(* IEC 61131-3 sources: plc-st-coding-agent/progress/evidence/f14_v8_temperature_repair_20261113/jobs/custom_deepseek-v4pro, 8 files *)

(* ---- public-medium-04.candidate_01.st ---- *)
FUNCTION_BLOCK FB_TemperatureControl
VAR_INPUT
    TemperatureSensorInput : REAL;
    SetTemperature : REAL;
END_VAR
VAR_OUTPUT
    CurrentTemperature : REAL;
    SetTempDisplay : REAL;
    HeaterStatus : BOOL;
    OverheatProtection : BOOL;
    HeaterOutput : BOOL;
END_VAR
VAR
    sensor_fault : BOOL;
    heater_request : BOOL;
    overheat_active : BOOL;
    tmp_heater_enable : BOOL;
    HeatingTimer : TON;
    CoolingTimer : TON;
END_VAR

(* ENGINEERING_CONTRACT
   O1 CurrentTemperature: copies TemperatureSensorInput; no fault suppression; units = input units (PUB006/PUB007).
   O2 SetTempDisplay: copies SetTemperature; units same as input (PUB006/PUB007).
   O3 HeaterStatus: copies final HeaterOutput; true while actual heater command active (PUB006/PUB007).
   O4 OverheatProtection: latched TRUE when heater has been continuously enabled for **strictly more than 5 s** (PUB005).
       Cleared automatically after a 3 s cooling period measured with CoolingTimer (PUB005).
       No external reset; state is retained during the 3 s cooldown.
   O5 HeaterOutput: TRUE when sensor input in [0,100] and TemperatureSensorInput < SetTemperature and not overheat-active (PUB003/PUB004/PUB005/PUB008).
       FALSE on sensor fault (input <0 or >100), on overheat, or when temperature >= setpoint.
   State retention: OverheatProtection held during 3 s wait; HeatingTimer resets whenever heater enable goes FALSE;
       CoolingTimer resets when overheat becomes inactive.
   Same‑scan priority: overheat trigger and heater disable occur in the same scan in which the strict >5 s condition is first satisfied;
       when cooling completes, heater may re‑enable in the same scan if the low‑temperature condition still holds.
   Boundaries: heater start condition is strict “<”; fault uses “<0.0 OR >100.0” (both exclusive); exact 0/100 are valid.
       TIMER thresholds use TIME constants; strict “>5 s” is implemented by requiring the 5 s threshold to have been reached in a previous scan
       and the heater still enabled in the current scan, thereby ensuring a positive elapsed time beyond 5 s.
*)
(* CONTRACT_RULES [] *)

// 1. Compute sensor fault and basic heater request
sensor_fault := (TemperatureSensorInput < 0.0) OR (TemperatureSensorInput > 100.0);
heater_request := NOT sensor_fault AND (TemperatureSensorInput < SetTemperature);

// 2. Determine heater enable before any new overheat decision (uses previous overheat state)
tmp_heater_enable := heater_request AND NOT overheat_active;

// 3. Detect strict overheat: HeatingTimer had already reached 5 s in the previous scan (Q true)
//    and the heater is still enabled now -> elapsed time > 5 s.
IF HeatingTimer.Q AND tmp_heater_enable THEN
    overheat_active := TRUE;
    tmp_heater_enable := FALSE;   // force heater off immediately in this scan
END_IF;

// 4. Update 5‑second timer with the current (possibly corrected) enable signal
HeatingTimer(IN := tmp_heater_enable, PT := T#5S);

// 5. Update cooling timer (3 s)
CoolingTimer(IN := overheat_active, PT := T#3S);
IF overheat_active AND CoolingTimer.Q THEN
    overheat_active := FALSE;      // cooling period finished, protection cleared
END_IF;

// 6. Final outputs
CurrentTemperature := TemperatureSensorInput;
SetTempDisplay := SetTemperature;
HeaterOutput := heater_request AND NOT overheat_active;
HeaterStatus := HeaterOutput;
OverheatProtection := overheat_active;

END_FUNCTION_BLOCK

(* ---- public-medium-04.candidate_02.st ---- *)
FUNCTION_BLOCK FB_TemperatureControl
VAR_INPUT
    TemperatureSensorInput : REAL;
    SetTemperature : REAL;
END_VAR
VAR_OUTPUT
    CurrentTemperature : REAL;
    SetTempDisplay : REAL;
    HeaterStatus : BOOL;
    OverheatProtection : BOOL;
    HeaterOutput : BOOL;
END_VAR
VAR
    sensor_fault : BOOL;
    heater_request : BOOL;
    overheat_active : BOOL;
    tmp_heater_enable : BOOL;
    HeatingTimer : TON;
    CoolingTimer : TON;
END_VAR

(* ENGINEERING_CONTRACT
   O1 CurrentTemperature: copies TemperatureSensorInput; no fault suppression; units = input units (PUB006/PUB007).
   O2 SetTempDisplay: copies SetTemperature; units same as input (PUB006/PUB007).
   O3 HeaterStatus: copies final HeaterOutput; true while actual heater command active (PUB006/PUB007).
   O4 OverheatProtection: latched TRUE when heater has been continuously enabled for at least 5 seconds (PUB005).
       Cleared automatically after a 3 second cooling period measured with CoolingTimer (PUB005).
       No external reset; state is retained during the 3 s cooldown.
   O5 HeaterOutput: TRUE when sensor input in [0,100] and TemperatureSensorInput < SetTemperature and not overheat-active
       (PUB003/PUB004/PUB005/PUB008). FALSE on sensor fault (input <0 or >100), on overheat, or when temperature >= setpoint.
   State retention: OverheatProtection held during 3 s wait; HeatingTimer resets whenever heater enable goes FALSE;
       CoolingTimer resets when overheat becomes inactive.
   Same‑scan priority: overheat trigger and heater disable occur in the same scan in which the 5 s threshold is reached;
       when cooling completes, heater may re‑enable in the same scan if the low‑temperature condition still holds.
   Boundaries: heater start condition is strict “<”; fault uses “<0.0 OR >100.0” (both exclusive); exact 0/100 are valid.
       TIMER thresholds use TIME constants; “≥5 s” for overheat and “≥3 s” for cooldown are implemented with standard TON.Q.
*)
(* CONTRACT_RULES [] *)

// 1. Compute sensor fault and basic heater request
sensor_fault := (TemperatureSensorInput < 0.0) OR (TemperatureSensorInput > 100.0);
heater_request := NOT sensor_fault AND (TemperatureSensorInput < SetTemperature);

// 2. Determine heater enable before overheat decision (uses previous overheat state)
tmp_heater_enable := heater_request AND NOT overheat_active;

// 3. Update 5‑second timer with current enable
HeatingTimer(IN := tmp_heater_enable, PT := T#5S);

// 4. Trigger overheat immediately when timer reaches PT (≥5 s)
IF HeatingTimer.Q AND tmp_heater_enable THEN
    overheat_active := TRUE;
END_IF;

// 5. Update cooling timer (3 s)
CoolingTimer(IN := overheat_active, PT := T#3S);

// 6. Clear overheat when cooling time reaches 3 s
IF overheat_active AND CoolingTimer.Q THEN
    overheat_active := FALSE;
END_IF;

// 7. Final outputs
CurrentTemperature := TemperatureSensorInput;
SetTempDisplay := SetTemperature;
HeaterOutput := heater_request AND NOT overheat_active;
HeaterStatus := HeaterOutput;
OverheatProtection := overheat_active;

END_FUNCTION_BLOCK

(* ---- public-medium-04.candidate_03.st ---- *)
FUNCTION_BLOCK FB_TemperatureControl
VAR_INPUT
    TemperatureSensorInput : REAL;
    SetTemperature : REAL;
END_VAR
VAR_OUTPUT
    CurrentTemperature : REAL;
    SetTempDisplay : REAL;
    HeaterStatus : BOOL;
    OverheatProtection : BOOL;
    HeaterOutput : BOOL;
END_VAR
VAR
    sensor_fault : BOOL;
    heater_request : BOOL;
    overheat_active : BOOL;
    tmp_heater_enable : BOOL;
    HeatingTimer : TON;
    CoolingTimer : TON;
END_VAR

(* ENGINEERING_CONTRACT
   O1 CurrentTemperature: copies TemperatureSensorInput; no fault suppression; units = input units (PUB006/PUB007).
   O2 SetTempDisplay: copies SetTemperature; units same as input (PUB006/PUB007).
   O3 HeaterStatus: copies final HeaterOutput; true while actual heater command active (PUB006/PUB007).
   O4 OverheatProtection: latched TRUE when heater has been continuously enabled for **strictly more than 5 seconds**
       (PUB005). HeatingTimer uses a large PT and compares ET > T#5S to enforce strict >.
       Cleared automatically after a 3 second cooling period: CoolingTimer.Q (ET >= T#3S).
       No external reset; state retained during cooldown.
   O5 HeaterOutput: TRUE when sensor input in [0,100] AND TemperatureSensorInput < SetTemperature AND NOT overheat_active
       (PUB003/PUB004/PUB005/PUB008). FALSE on sensor fault, overheat, or temp >= setpoint.
   State retention: OverheatProtection held during 3 s wait; HeatingTimer resets whenever heater enable goes FALSE;
       CoolingTimer resets when overheat becomes inactive.
   Same‑scan priority: overheat trigger and heater disable occur in the same scan when ET > 5 s is detected.
       When cooling completes, heater may re‑enable in the same scan if low‑temperature condition still holds.
   Boundaries: heater start condition is strict “<”; fault uses “<0.0 OR >100.0” (exclusive); exact 0/100 are valid.
       Overheat uses “>5 s”; cooldown uses “>=3 s”.
*)
(* CONTRACT_RULES [] *)

// 1. Compute sensor fault and basic heater request
sensor_fault := (TemperatureSensorInput < 0.0) OR (TemperatureSensorInput > 100.0);
heater_request := NOT sensor_fault AND (TemperatureSensorInput < SetTemperature);

// 2. Determine heater enable before overheat decision (uses previous overheat state)
tmp_heater_enable := heater_request AND NOT overheat_active;

// 3. Update heating timer with a large PT so ET can exceed T#5S
HeatingTimer(IN := tmp_heater_enable, PT := T#1D);
IF tmp_heater_enable AND (HeatingTimer.ET > T#5S) THEN
    overheat_active := TRUE;
END_IF;

// 4. Update cooling timer (standard TON: Q becomes TRUE at >= T#3S)
CoolingTimer(IN := overheat_active, PT := T#3S);
IF overheat_active AND CoolingTimer.Q THEN
    overheat_active := FALSE;
END_IF;

// 5. Final outputs
CurrentTemperature := TemperatureSensorInput;
SetTempDisplay := SetTemperature;
HeaterOutput := heater_request AND NOT overheat_active;
HeaterStatus := HeaterOutput;
OverheatProtection := overheat_active;

END_FUNCTION_BLOCK

(* ---- public-medium-04.candidate_04.st ---- *)
FUNCTION_BLOCK FB_TemperatureControl
VAR_INPUT
    TemperatureSensorInput : REAL;
    SetTemperature : REAL;
END_VAR
VAR_OUTPUT
    CurrentTemperature : REAL;
    SetTempDisplay : REAL;
    HeaterStatus : BOOL;
    OverheatProtection : BOOL;
    HeaterOutput : BOOL;
END_VAR
VAR
    sensor_fault : BOOL;
    heater_request : BOOL;
    overheat_active : BOOL;
    local_heater_enable : BOOL;

    (* Free-running clock for measuring scan intervals *)
    ClockTimer : TON;
    prev_clock_et : TIME := T#0ms;

    (* Custom heating accumulator for strict >5s detection *)
    heater_on_accum : TIME := T#0ms;

    (* Cooling timer with standard TON (Q at >=3s) *)
    CoolingTimer : TON;
END_VAR

(* ENGINEERING_CONTRACT
   O1 CurrentTemperature: copies TemperatureSensorInput; no fault suppression; units = input units (PUB006/PUB007).
   O2 SetTempDisplay: copies SetTemperature; units same as input (PUB006/PUB007).
   O3 HeaterStatus: copies final HeaterOutput; true while actual heater command active (PUB006/PUB007).
   O4 OverheatProtection: latched TRUE when heater has been continuously enabled for **strictly more than 5 seconds**
       (PUB005). Uses custom TIME accumulator based on free-running TON delta to correctly include the
       first scan interval after enable. Cleared automatically after 3 s cooling: CoolingTimer.Q (ET >= T#3S).
       No external reset; state retained during cooldown.
   O5 HeaterOutput: TRUE when sensor input in [0,100] AND TemperatureSensorInput < SetTemperature AND NOT overheat_active
       (PUB003/PUB004/PUB005/PUB008). FALSE on sensor fault, overheat, or temp >= setpoint.
   State retention: OverheatProtection held during 3 s wait; heating accumulator resets when heater enable goes FALSE;
       CoolingTimer resets when overheat becomes inactive.
   Same-scan priority: overheat trigger and heater disable occur in the same scan when accumulated
       heater-on time exceeds 5 s. When cooling completes, heater may re-enable in the same scan if low-temperature
       condition still holds.
   Boundaries: heater start condition is strict “<”; fault uses “<0.0 OR >100.0” (exclusive); exact 0/100 are valid.
       Overheat uses “>5 s”; cooldown uses “>=3 s”. All TIME arithmetic is non-capped because ClockTimer PT is T#1D.
*)
(* CONTRACT_RULES [] *)

// 1. Compute sensor fault and basic heater request
sensor_fault := (TemperatureSensorInput < 0.0) OR (TemperatureSensorInput > 100.0);
heater_request := NOT sensor_fault AND (TemperatureSensorInput < SetTemperature);

// 2. Free-running clock for scan interval measurement
ClockTimer(IN := TRUE, PT := T#1D);
tmp_delta := ClockTimer.ET - prev_clock_et;
prev_clock_et := ClockTimer.ET;

// 3. Heater enable before overheat decision (uses previous overheat state)
local_heater_enable := heater_request AND NOT overheat_active;

// 4. Update heating accumulator (measures continuous heater-on time, including current scan)
IF local_heater_enable THEN
    heater_on_accum := heater_on_accum + tmp_delta;
ELSE
    heater_on_accum := T#0ms;
END_IF;

// 5. Overheat protection trigger: strictly more than 5 s
IF heater_on_accum > T#5S THEN
    overheat_active := TRUE;
END_IF;

// 6. Cooling timer (standard TON; clears after 3 s)
CoolingTimer(IN := overheat_active, PT := T#3S);
IF overheat_active AND CoolingTimer.Q THEN
    overheat_active := FALSE;
END_IF;

// 7. Final outputs
CurrentTemperature := TemperatureSensorInput;
SetTempDisplay := SetTemperature;
HeaterOutput := heater_request AND NOT overheat_active;
HeaterStatus := HeaterOutput;
OverheatProtection := overheat_active;

END_FUNCTION_BLOCK

(* ---- public-medium-04.raw_candidate_01.st ---- *)
FUNCTION_BLOCK FB_TemperatureControl
VAR_INPUT
    TemperatureSensorInput : REAL;
    SetTemperature : REAL;
END_VAR
VAR_OUTPUT
    CurrentTemperature : REAL;
    SetTempDisplay : REAL;
    HeaterStatus : BOOL;
    OverheatProtection : BOOL;
    HeaterOutput : BOOL;
END_VAR
VAR
    sensor_fault : BOOL;
    heater_request : BOOL;
    overheat_active : BOOL;
    tmp_heater_enable : BOOL;
    HeatingTimer : TON;
    CoolingTimer : TON;
END_VAR

(* ENGINEERING_CONTRACT
   O1 CurrentTemperature: copies TemperatureSensorInput; no fault suppression; units = input units (PUB006/PUB007).
   O2 SetTempDisplay: copies SetTemperature; units same as input (PUB006/PUB007).
   O3 HeaterStatus: copies final HeaterOutput; true while actual heater command active (PUB006/PUB007).
   O4 OverheatProtection: latched TRUE when heater has been continuously enabled for **strictly more than 5 s** (PUB005).
       Cleared automatically after a 3 s cooling period measured with CoolingTimer (PUB005).
       No external reset; state is retained during the 3 s cooldown.
   O5 HeaterOutput: TRUE when sensor input in [0,100] and TemperatureSensorInput < SetTemperature and not overheat-active (PUB003/PUB004/PUB005/PUB008).
       FALSE on sensor fault (input <0 or >100), on overheat, or when temperature >= setpoint.
   State retention: OverheatProtection held during 3 s wait; HeatingTimer resets whenever heater enable goes FALSE;
       CoolingTimer resets when overheat becomes inactive.
   Same‑scan priority: overheat trigger and heater disable occur in the same scan in which the strict >5 s condition is first satisfied;
       when cooling completes, heater may re‑enable in the same scan if the low‑temperature condition still holds.
   Boundaries: heater start condition is strict “<”; fault uses “<0.0 OR >100.0” (both exclusive); exact 0/100 are valid.
       TIMER thresholds use TIME constants; strict “>5 s” is implemented by requiring the 5 s threshold to have been reached in a previous scan
       and the heater still enabled in the current scan, thereby ensuring a positive elapsed time beyond 5 s.
*)
(* CONTRACT_RULES [] *)

// 1. Compute sensor fault and basic heater request
sensor_fault := (TemperatureSensorInput < 0.0) OR (TemperatureSensorInput > 100.0);
heater_request := NOT sensor_fault AND (TemperatureSensorInput < SetTemperature);

// 2. Determine heater enable before any new overheat decision (uses previous overheat state)
tmp_heater_enable := heater_request AND NOT overheat_active;

// 3. Detect strict overheat: HeatingTimer had already reached 5 s in the previous scan (Q true)
//    and the heater is still enabled now -> elapsed time > 5 s.
IF HeatingTimer.Q AND tmp_heater_enable THEN
    overheat_active := TRUE;
    tmp_heater_enable := FALSE;   // force heater off immediately in this scan
END_IF;

// 4. Update 5‑second timer with the current (possibly corrected) enable signal
HeatingTimer(IN := tmp_heater_enable, PT := T#5S);

// 5. Update cooling timer (3 s)
CoolingTimer(IN := overheat_active, PT := T#3S);
IF overheat_active AND CoolingTimer.Q THEN
    overheat_active := FALSE;      // cooling period finished, protection cleared
END_IF;

// 6. Final outputs
CurrentTemperature := TemperatureSensorInput;
SetTempDisplay := SetTemperature;
HeaterOutput := heater_request AND NOT overheat_active;
HeaterStatus := HeaterOutput;
OverheatProtection := overheat_active;

END_FUNCTION_BLOCK

(* ---- public-medium-04.raw_candidate_02.st ---- *)
FUNCTION_BLOCK FB_TemperatureControl
VAR_INPUT
    TemperatureSensorInput : REAL;
    SetTemperature : REAL;
END_VAR
VAR_OUTPUT
    CurrentTemperature : REAL;
    SetTempDisplay : REAL;
    HeaterStatus : BOOL;
    OverheatProtection : BOOL;
    HeaterOutput : BOOL;
END_VAR
VAR
    sensor_fault : BOOL;
    heater_request : BOOL;
    overheat_active : BOOL;
    tmp_heater_enable : BOOL;
    HeatingTimer : TON;
    CoolingTimer : TON;
END_VAR

(* ENGINEERING_CONTRACT
   O1 CurrentTemperature: copies TemperatureSensorInput; no fault suppression; units = input units (PUB006/PUB007).
   O2 SetTempDisplay: copies SetTemperature; units same as input (PUB006/PUB007).
   O3 HeaterStatus: copies final HeaterOutput; true while actual heater command active (PUB006/PUB007).
   O4 OverheatProtection: latched TRUE when heater has been continuously enabled for at least 5 seconds (PUB005).
       Cleared automatically after a 3 second cooling period measured with CoolingTimer (PUB005).
       No external reset; state is retained during the 3 s cooldown.
   O5 HeaterOutput: TRUE when sensor input in [0,100] and TemperatureSensorInput < SetTemperature and not overheat-active
       (PUB003/PUB004/PUB005/PUB008). FALSE on sensor fault (input <0 or >100), on overheat, or when temperature >= setpoint.
   State retention: OverheatProtection held during 3 s wait; HeatingTimer resets whenever heater enable goes FALSE;
       CoolingTimer resets when overheat becomes inactive.
   Same‑scan priority: overheat trigger and heater disable occur in the same scan in which the 5 s threshold is reached;
       when cooling completes, heater may re‑enable in the same scan if the low‑temperature condition still holds.
   Boundaries: heater start condition is strict “<”; fault uses “<0.0 OR >100.0” (both exclusive); exact 0/100 are valid.
       TIMER thresholds use TIME constants; “≥5 s” for overheat and “≥3 s” for cooldown are implemented with standard TON.Q.
*)
(* CONTRACT_RULES [] *)

// 1. Compute sensor fault and basic heater request
sensor_fault := (TemperatureSensorInput < 0.0) OR (TemperatureSensorInput > 100.0);
heater_request := NOT sensor_fault AND (TemperatureSensorInput < SetTemperature);

// 2. Determine heater enable before overheat decision (uses previous overheat state)
tmp_heater_enable := heater_request AND NOT overheat_active;

// 3. Update 5‑second timer with current enable
HeatingTimer(IN := tmp_heater_enable, PT := T#5S);

// 4. Trigger overheat immediately when timer reaches PT (≥5 s)
IF HeatingTimer.Q AND tmp_heater_enable THEN
    overheat_active := TRUE;
END_IF;

// 5. Update cooling timer (3 s)
CoolingTimer(IN := overheat_active, PT := T#3S);

// 6. Clear overheat when cooling time reaches 3 s
IF overheat_active AND CoolingTimer.Q THEN
    overheat_active := FALSE;
END_IF;

// 7. Final outputs
CurrentTemperature := TemperatureSensorInput;
SetTempDisplay := SetTemperature;
HeaterOutput := heater_request AND NOT overheat_active;
HeaterStatus := HeaterOutput;
OverheatProtection := overheat_active;

END_FUNCTION_BLOCK

(* ---- public-medium-04.raw_candidate_03.st ---- *)
FUNCTION_BLOCK FB_TemperatureControl
VAR_INPUT
    TemperatureSensorInput : REAL;
    SetTemperature : REAL;
END_VAR
VAR_OUTPUT
    CurrentTemperature : REAL;
    SetTempDisplay : REAL;
    HeaterStatus : BOOL;
    OverheatProtection : BOOL;
    HeaterOutput : BOOL;
END_VAR
VAR
    sensor_fault : BOOL;
    heater_request : BOOL;
    overheat_active : BOOL;
    tmp_heater_enable : BOOL;
    HeatingTimer : TON;
    CoolingTimer : TON;
END_VAR

(* ENGINEERING_CONTRACT
   O1 CurrentTemperature: copies TemperatureSensorInput; no fault suppression; units = input units (PUB006/PUB007).
   O2 SetTempDisplay: copies SetTemperature; units same as input (PUB006/PUB007).
   O3 HeaterStatus: copies final HeaterOutput; true while actual heater command active (PUB006/PUB007).
   O4 OverheatProtection: latched TRUE when heater has been continuously enabled for **strictly more than 5 seconds**
       (PUB005). HeatingTimer uses a large PT and compares ET > T#5S to enforce strict >.
       Cleared automatically after a 3 second cooling period: CoolingTimer.Q (ET >= T#3S).
       No external reset; state retained during cooldown.
   O5 HeaterOutput: TRUE when sensor input in [0,100] AND TemperatureSensorInput < SetTemperature AND NOT overheat_active
       (PUB003/PUB004/PUB005/PUB008). FALSE on sensor fault, overheat, or temp >= setpoint.
   State retention: OverheatProtection held during 3 s wait; HeatingTimer resets whenever heater enable goes FALSE;
       CoolingTimer resets when overheat becomes inactive.
   Same‑scan priority: overheat trigger and heater disable occur in the same scan when ET > 5 s is detected.
       When cooling completes, heater may re‑enable in the same scan if low‑temperature condition still holds.
   Boundaries: heater start condition is strict “<”; fault uses “<0.0 OR >100.0” (exclusive); exact 0/100 are valid.
       Overheat uses “>5 s”; cooldown uses “>=3 s”.
*)
(* CONTRACT_RULES [] *)

// 1. Compute sensor fault and basic heater request
sensor_fault := (TemperatureSensorInput < 0.0) OR (TemperatureSensorInput > 100.0);
heater_request := NOT sensor_fault AND (TemperatureSensorInput < SetTemperature);

// 2. Determine heater enable before overheat decision (uses previous overheat state)
tmp_heater_enable := heater_request AND NOT overheat_active;

// 3. Update heating timer with a large PT so ET can exceed T#5S
HeatingTimer(IN := tmp_heater_enable, PT := T#1D);
IF tmp_heater_enable AND (HeatingTimer.ET > T#5S) THEN
    overheat_active := TRUE;
END_IF;

// 4. Update cooling timer (standard TON: Q becomes TRUE at >= T#3S)
CoolingTimer(IN := overheat_active, PT := T#3S);
IF overheat_active AND CoolingTimer.Q THEN
    overheat_active := FALSE;
END_IF;

// 5. Final outputs
CurrentTemperature := TemperatureSensorInput;
SetTempDisplay := SetTemperature;
HeaterOutput := heater_request AND NOT overheat_active;
HeaterStatus := HeaterOutput;
OverheatProtection := overheat_active;

END_FUNCTION_BLOCK

(* ---- public-medium-04.raw_candidate_04.st ---- *)
FUNCTION_BLOCK FB_TemperatureControl
VAR_INPUT
    TemperatureSensorInput : REAL;
    SetTemperature : REAL;
END_VAR
VAR_OUTPUT
    CurrentTemperature : REAL;
    SetTempDisplay : REAL;
    HeaterStatus : BOOL;
    OverheatProtection : BOOL;
    HeaterOutput : BOOL;
END_VAR
VAR
    sensor_fault : BOOL;
    heater_request : BOOL;
    overheat_active : BOOL;
    local_heater_enable : BOOL;

    (* Free-running clock for measuring scan intervals *)
    ClockTimer : TON;
    prev_clock_et : TIME := T#0ms;

    (* Custom heating accumulator for strict >5s detection *)
    heater_on_accum : TIME := T#0ms;

    (* Cooling timer with standard TON (Q at >=3s) *)
    CoolingTimer : TON;
END_VAR

(* ENGINEERING_CONTRACT
   O1 CurrentTemperature: copies TemperatureSensorInput; no fault suppression; units = input units (PUB006/PUB007).
   O2 SetTempDisplay: copies SetTemperature; units same as input (PUB006/PUB007).
   O3 HeaterStatus: copies final HeaterOutput; true while actual heater command active (PUB006/PUB007).
   O4 OverheatProtection: latched TRUE when heater has been continuously enabled for **strictly more than 5 seconds**
       (PUB005). Uses custom TIME accumulator based on free-running TON delta to correctly include the
       first scan interval after enable. Cleared automatically after 3 s cooling: CoolingTimer.Q (ET >= T#3S).
       No external reset; state retained during cooldown.
   O5 HeaterOutput: TRUE when sensor input in [0,100] AND TemperatureSensorInput < SetTemperature AND NOT overheat_active
       (PUB003/PUB004/PUB005/PUB008). FALSE on sensor fault, overheat, or temp >= setpoint.
   State retention: OverheatProtection held during 3 s wait; heating accumulator resets when heater enable goes FALSE;
       CoolingTimer resets when overheat becomes inactive.
   Same-scan priority: overheat trigger and heater disable occur in the same scan when accumulated
       heater-on time exceeds 5 s. When cooling completes, heater may re-enable in the same scan if low-temperature
       condition still holds.
   Boundaries: heater start condition is strict “<”; fault uses “<0.0 OR >100.0” (exclusive); exact 0/100 are valid.
       Overheat uses “>5 s”; cooldown uses “>=3 s”. All TIME arithmetic is non-capped because ClockTimer PT is T#1D.
*)
(* CONTRACT_RULES [] *)

// 1. Compute sensor fault and basic heater request
sensor_fault := (TemperatureSensorInput < 0.0) OR (TemperatureSensorInput > 100.0);
heater_request := NOT sensor_fault AND (TemperatureSensorInput < SetTemperature);

// 2. Free-running clock for scan interval measurement
ClockTimer(IN := TRUE, PT := T#1D);
tmp_delta := ClockTimer.ET - prev_clock_et;
prev_clock_et := ClockTimer.ET;

// 3. Heater enable before overheat decision (uses previous overheat state)
local_heater_enable := heater_request AND NOT overheat_active;

// 4. Update heating accumulator (measures continuous heater-on time, including current scan)
IF local_heater_enable THEN
    heater_on_accum := heater_on_accum + tmp_delta;
ELSE
    heater_on_accum := T#0ms;
END_IF;

// 5. Overheat protection trigger: strictly more than 5 s
IF heater_on_accum > T#5S THEN
    overheat_active := TRUE;
END_IF;

// 6. Cooling timer (standard TON; clears after 3 s)
CoolingTimer(IN := overheat_active, PT := T#3S);
IF overheat_active AND CoolingTimer.Q THEN
    overheat_active := FALSE;
END_IF;

// 7. Final outputs
CurrentTemperature := TemperatureSensorInput;
SetTempDisplay := SetTemperature;
HeaterOutput := heater_request AND NOT overheat_active;
HeaterStatus := HeaterOutput;
OverheatProtection := overheat_active;

END_FUNCTION_BLOCK
